(* Logix 5000 project; controller TFF vendor 1 type 14 code 107 rev 33.11; software revision 33.04; part 32 of 38 *)
(* tags used below, declared in another part *)
   ModbusLogTimer : TIMER;
   TIME : DINT[2];
   TimeInSecondsDINT : DINT;
   AI101 : ALIAS FOR AnalogPoint[16];
   AI202 : ALIAS FOR AnalogPoint[9];
   AP008 : ALIAS FOR DigitalOutput[14];
   ARC_AI101 : ARC_pH;
   ARC_AI202 : ARC_pH;
   BagInflate : BagInflate;
   DPAlarm : ALIAS FOR AlarmAnalog[40];
   FlowPath : FlowPath[64];   // Flow Path Array
   GWModbus : IO_Station;   // Status of Gateway Modbus
   IBA001 : ALIAS FOR DigitalOutput[25];
   Membrane_Data : Membrane_Data;   // Membrane Data
   ModbusTimeSyncTimer : TIMER;
   OperatingTime : OperatingTime;
   Options : Options;   // Options List
   Phase0 : ALIAS FOR Phase[0];   // Phase 0
   PI601 : ALIAS FOR AnalogPoint[21];
   PipeAnimation : PipeAnimation;   // HMI Pipe Animation Array
   SIC001_AO : ALIAS FOR AnalogOutput[0];
   SIC001_DO : ALIAS FOR DigitalOutput[8];
   SIC002_AO : ALIAS FOR AnalogOutput[1];
   SIC002_DO : ALIAS FOR DigitalOutput[9];
   SysControl : SysControl;   // General system status and command
   TimerControl : TimerControl;   // Timer Control
   TMPAlarm : ALIAS FOR AlarmAnalog[41];
   YA41 : ALIAS FOR DigitalPoint[73];
(* Process, continued *)

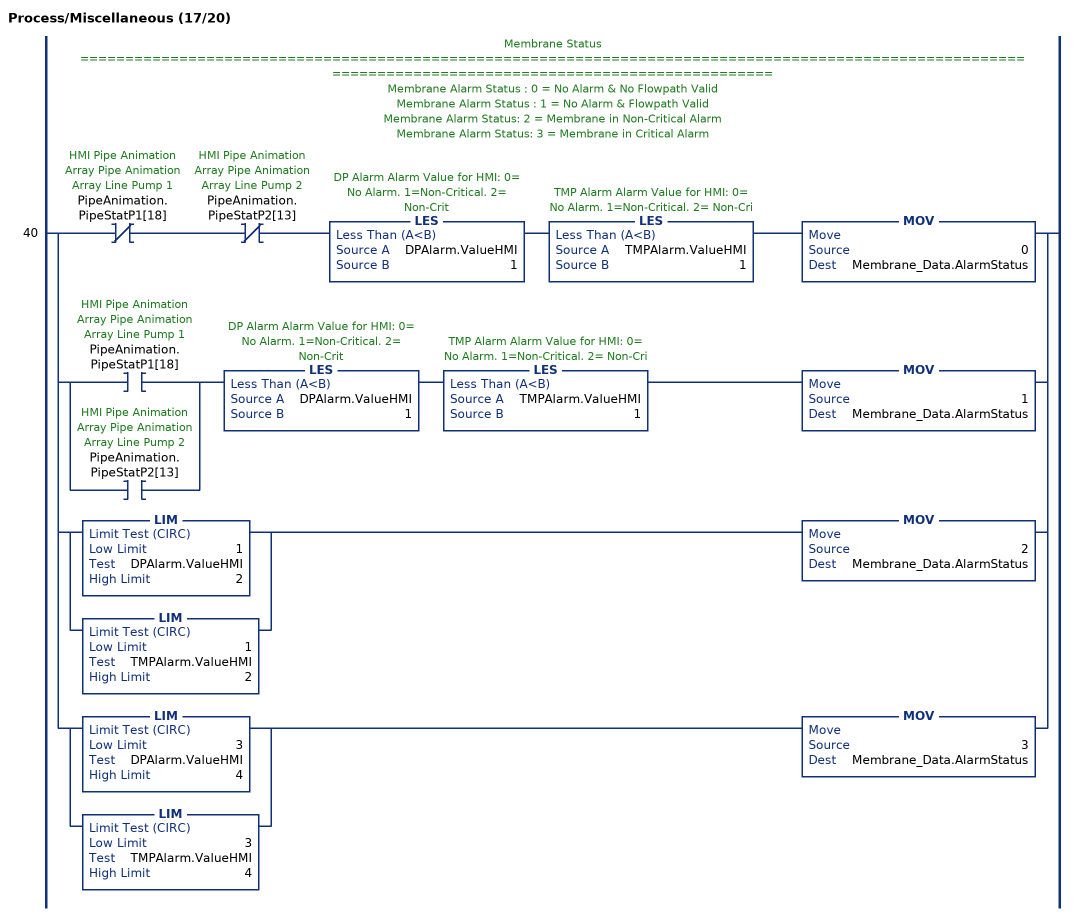
   [picture p374: Process/Miscellaneous rungs 40-40]
   // Membrane Status
   // ==========================================================================================================================================================
   // Membrane Alarm Status : 0 = No Alarm & No Flowpath Valid
   // Membrane Alarm Status : 1 = No Alarm & Flowpath Valid
   // Membrane Alarm Status: 2 = Membrane in Non-Critical Alarm
   // Membrane Alarm Status: 3 = Membrane in Critical Alarm
   40: [XIO(PipeAnimation.PipeStatP1[18]) XIO(PipeAnimation.PipeStatP2[13]) LES(DPAlarm.ValueHMI,1) LES(TMPAlarm.ValueHMI,1) MOV(0,Membrane_Data.AlarmStatus) ,[XIC(PipeAnimation.PipeStatP1[18]) ,XIC(PipeAnimation.PipeStatP2[13]) ] LES(DPAlarm.ValueHMI,1) LES(TMPAlarm.ValueHMI,1) MOV(1,Membrane_Data.AlarmStatus) ,[LIM(1,DPAlarm.ValueHMI,2) ,LIM(1,TMPAlarm.ValueHMI,2) ] MOV(2,Membrane_Data.AlarmStatus) ,[LIM(3,DPAlarm.ValueHMI,4) ,LIM(3,TMPAlarm.ValueHMI,4) ] MOV(3,Membrane_Data.AlarmStatus) ];
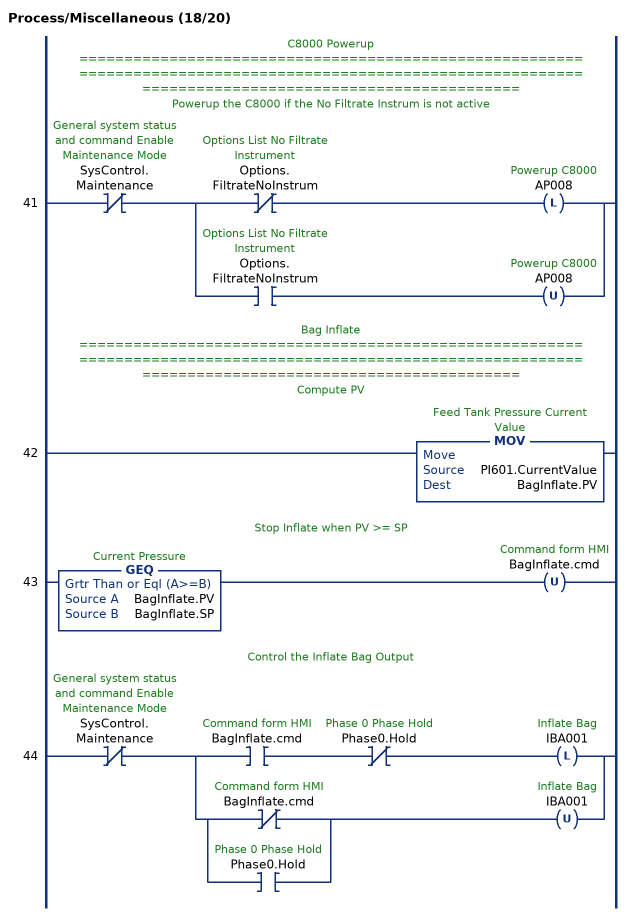
   // C8000 Powerup
   // ==========================================================================================================================================================
   // Powerup the C8000 if the No Filtrate Instrum is not active
   41: XIO(SysControl.Maintenance)[XIO(Options.FiltrateNoInstrum) OTL(AP008) ,XIC(Options.FiltrateNoInstrum) OTU(AP008) ];
   // Bag Inflate
   // ==========================================================================================================================================================
   // Compute PV
   42: MOV(PI601.CurrentValue,BagInflate.PV);
   // Stop Inflate when PV >= SP
   43: GEQ(BagInflate.PV,BagInflate.SP)OTU(BagInflate.cmd);
   // Control the Inflate Bag Output
   44: XIO(SysControl.Maintenance)[XIC(BagInflate.cmd) XIO(Phase0.Hold) OTL(IBA001) ,[XIO(BagInflate.cmd) ,XIC(Phase0.Hold) ] OTU(IBA001) ];
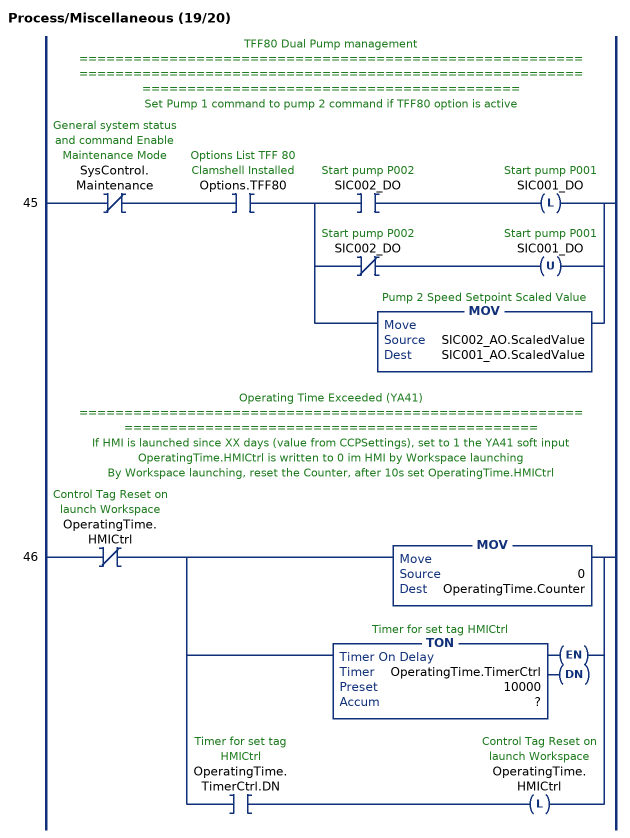
   // TFF80 Dual Pump management
   // ==========================================================================================================================================================
   // Set Pump 1 command to pump 2 command if TFF80 option is active
   45: XIO(SysControl.Maintenance)XIC(Options.TFF80)[[XIC(SIC002_DO) OTL(SIC001_DO) ,XIO(SIC002_DO) OTU(SIC001_DO) ] ,MOV(SIC002_AO.ScaledValue,SIC001_AO.ScaledValue) ];
   // Operating Time Exceeded (YA41)
   // ======================================================================================================
   // If HMI is launched since XX days (value from CCPSettings), set to 1 the YA41 soft input
   // OperatingTime.HMICtrl is written to 0 im HMI by Workspace launching
   // By Workspace launching, reset the Counter, after 10s set OperatingTime.HMICtrl
   46: XIO(OperatingTime.HMICtrl)[MOV(0,OperatingTime.Counter) ,TON(OperatingTime.TimerCtrl,?,?) ,XIC(OperatingTime.TimerCtrl.DN) OTL(OperatingTime.HMICtrl) ];
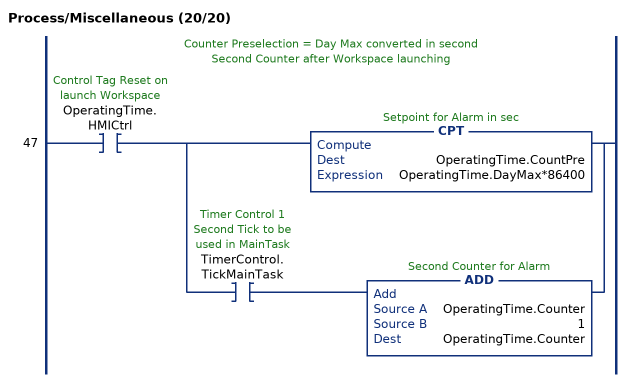
   // Counter Preselection = Day Max converted in second
   // Second Counter after Workspace launching
   47: XIC(OperatingTime.HMICtrl)[CPT(OperatingTime.CountPre,OperatingTime.DayMax*86400) ,XIC(TimerControl.TickMainTask) ADD(OperatingTime.Counter,1,OperatingTime.Counter) ];
END_ROUTINE

ROUTINE ModbusGateway   (* ladder *)
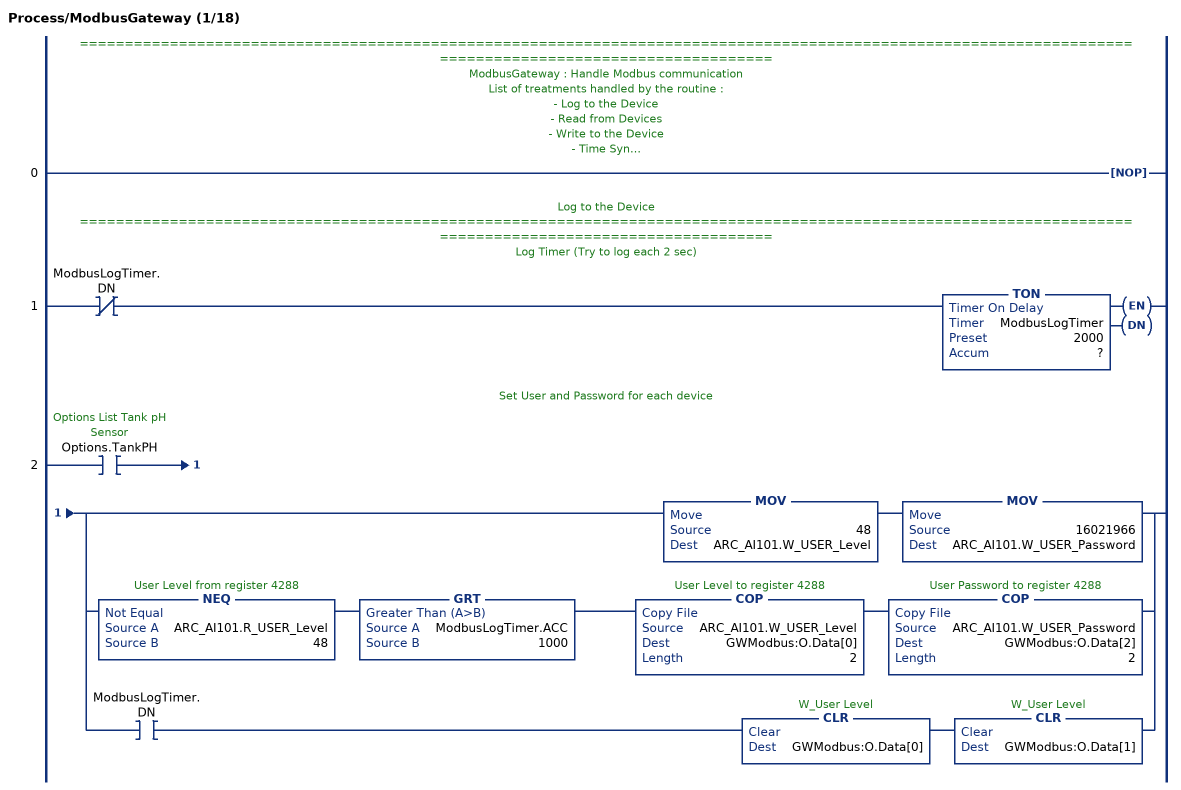
   // ==========================================================================================================================================================
   //                                                                                                                                 ModbusGateway : Handle Modbus communication
   //                                                     List of treatments handled by the routine :
   //                                                         - Log to the Device
   //                                                          - Read from Devices
   //                                                          - Write to the Device
   //                                                        - Time Sync
   //                                                     -----------------------------------------------------------------------------------------------------------------------------------------------------
   //                                                     History
   // 		2019-DEC-24 - Merck - Q. Spindler - Initial version for Candidate Release 1.00.00.00.a
   // ==========================================================================================================================================================
   0: NOP();
   // Log to the Device
   // ==========================================================================================================================================================
   // Log Timer (Try to log each 2 sec)
   1: XIO(ModbusLogTimer.DN)TON(ModbusLogTimer,?,?);
   // Set User and Password for each device
   2: XIC(Options.TankPH)[MOV(48,ARC_AI101.W_USER_Level) MOV(16021966,ARC_AI101.W_USER_Password) ,NEQ(ARC_AI101.R_USER_Level,48) GRT(ModbusLogTimer.ACC,1000) COP(ARC_AI101.W_USER_Level,GWModbus:O.Data[0],2) COP(ARC_AI101.W_USER_Password,GWModbus:O.Data[2],2) ,XIC(ModbusLogTimer.DN) CLR(GWModbus:O.Data[0]) CLR(GWModbus:O.Data[1]) ];
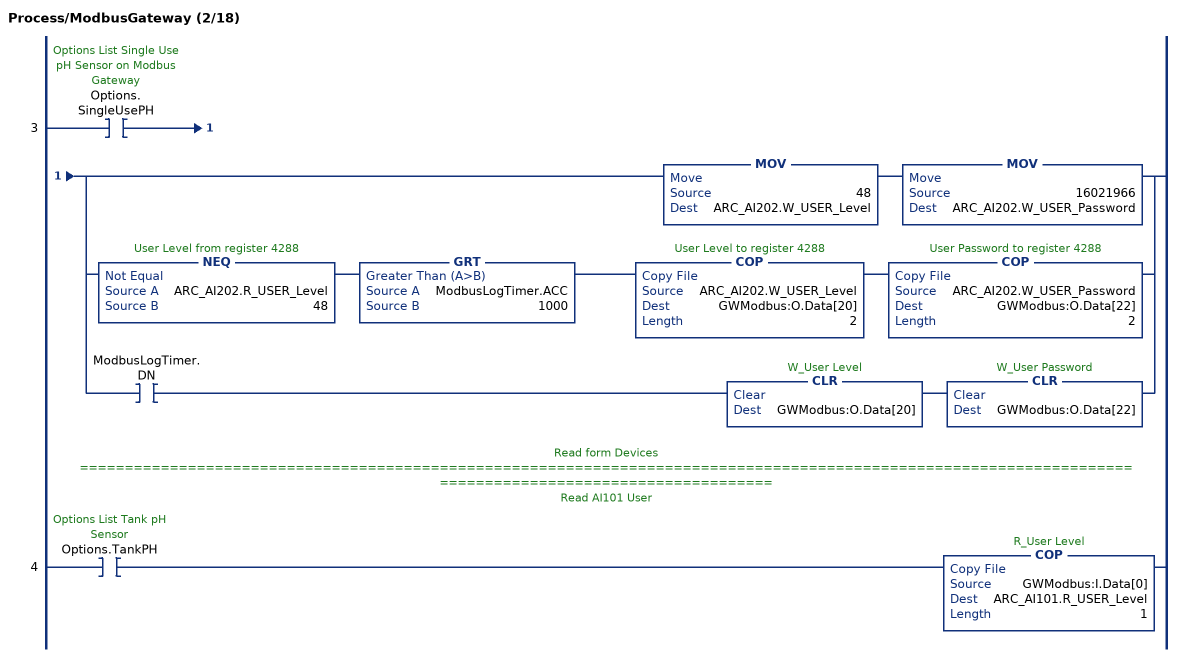
   3: XIC(Options.SingleUsePH)[MOV(48,ARC_AI202.W_USER_Level) MOV(16021966,ARC_AI202.W_USER_Password) ,NEQ(ARC_AI202.R_USER_Level,48) GRT(ModbusLogTimer.ACC,1000) COP(ARC_AI202.W_USER_Level,GWModbus:O.Data[20],2) COP(ARC_AI202.W_USER_Password,GWModbus:O.Data[22],2) ,XIC(ModbusLogTimer.DN) CLR(GWModbus:O.Data[20]) CLR(GWModbus:O.Data[22]) ];
   // Read form Devices
   // ==========================================================================================================================================================
   // Read AI101 User
   4: XIC(Options.TankPH)COP(GWModbus:I.Data[0],ARC_AI101.R_USER_Level,1);
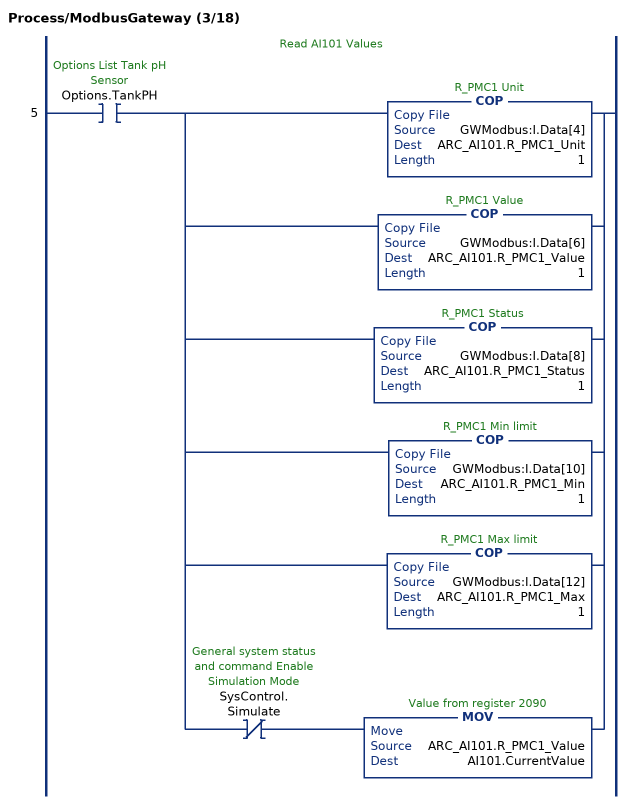
   // Read AI101 Values
   5: XIC(Options.TankPH)[COP(GWModbus:I.Data[4],ARC_AI101.R_PMC1_Unit,1) ,COP(GWModbus:I.Data[6],ARC_AI101.R_PMC1_Value,1) ,COP(GWModbus:I.Data[8],ARC_AI101.R_PMC1_Status,1) ,COP(GWModbus:I.Data[10],ARC_AI101.R_PMC1_Min,1) ,COP(GWModbus:I.Data[12],ARC_AI101.R_PMC1_Max,1) ,XIO(SysControl.Simulate) MOV(ARC_AI101.R_PMC1_Value,AI101.CurrentValue) ];
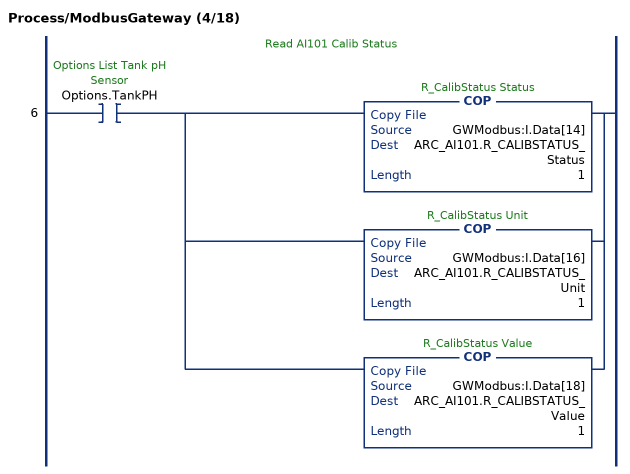
   // Read AI101 Calib Status
   6: XIC(Options.TankPH)[COP(GWModbus:I.Data[14],ARC_AI101.R_CALIBSTATUS_Status,1) ,COP(GWModbus:I.Data[16],ARC_AI101.R_CALIBSTATUS_Unit,1) ,COP(GWModbus:I.Data[18],ARC_AI101.R_CALIBSTATUS_Value,1) ];
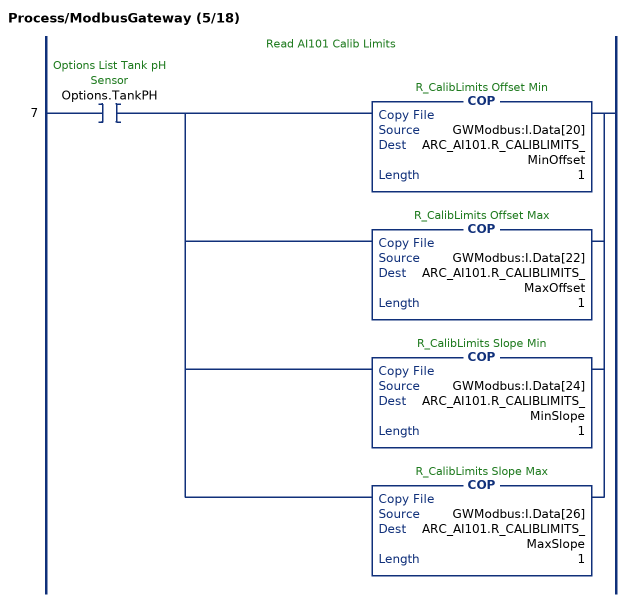
   // Read AI101 Calib Limits
   7: XIC(Options.TankPH)[COP(GWModbus:I.Data[20],ARC_AI101.R_CALIBLIMITS_MinOffset,1) ,COP(GWModbus:I.Data[22],ARC_AI101.R_CALIBLIMITS_MaxOffset,1) ,COP(GWModbus:I.Data[24],ARC_AI101.R_CALIBLIMITS_MinSlope,1) ,COP(GWModbus:I.Data[26],ARC_AI101.R_CALIBLIMITS_MaxSlope,1) ];
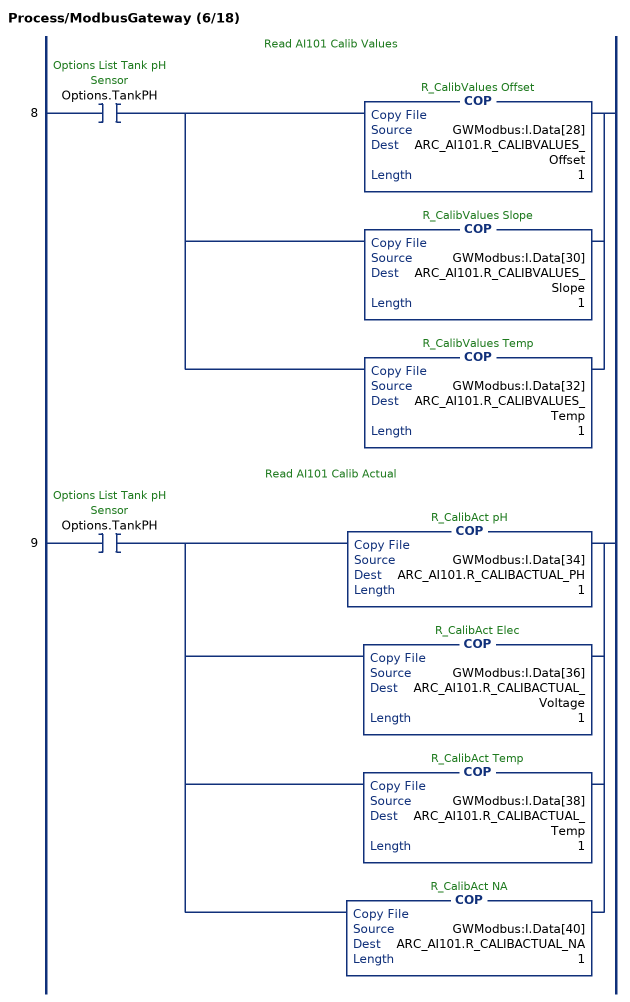
   // Read AI101 Calib Values
   8: XIC(Options.TankPH)[COP(GWModbus:I.Data[28],ARC_AI101.R_CALIBVALUES_Offset,1) ,COP(GWModbus:I.Data[30],ARC_AI101.R_CALIBVALUES_Slope,1) ,COP(GWModbus:I.Data[32],ARC_AI101.R_CALIBVALUES_Temp,1) ];
   // Read AI101 Calib Actual
   9: XIC(Options.TankPH)[COP(GWModbus:I.Data[34],ARC_AI101.R_CALIBACTUAL_PH,1) ,COP(GWModbus:I.Data[36],ARC_AI101.R_CALIBACTUAL_Voltage,1) ,COP(GWModbus:I.Data[38],ARC_AI101.R_CALIBACTUAL_Temp,1) ,COP(GWModbus:I.Data[40],ARC_AI101.R_CALIBACTUAL_NA,1) ];
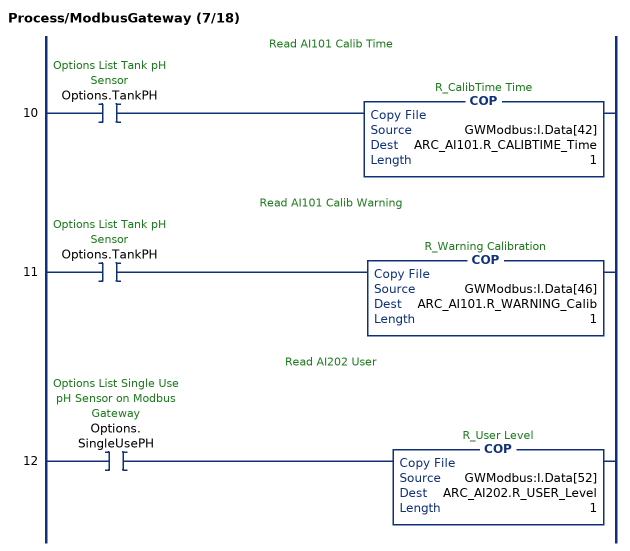
   // Read AI101 Calib Time
   10: XIC(Options.TankPH)COP(GWModbus:I.Data[42],ARC_AI101.R_CALIBTIME_Time,1);
   // Read AI101 Calib Warning
   11: XIC(Options.TankPH)COP(GWModbus:I.Data[46],ARC_AI101.R_WARNING_Calib,1);
   // Read AI202 User
   12: XIC(Options.SingleUsePH)COP(GWModbus:I.Data[52],ARC_AI202.R_USER_Level,1);
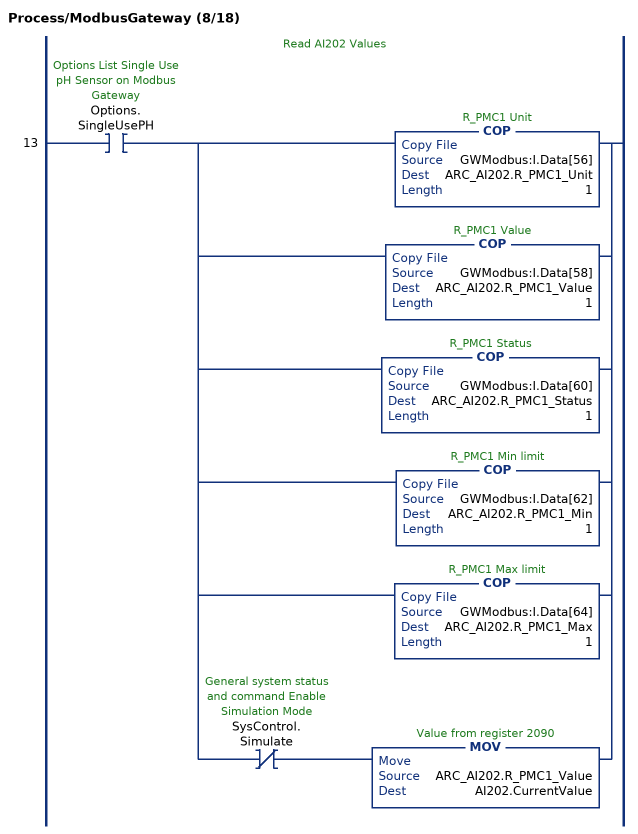
   // Read AI202 Values
   13: XIC(Options.SingleUsePH)[COP(GWModbus:I.Data[56],ARC_AI202.R_PMC1_Unit,1) ,COP(GWModbus:I.Data[58],ARC_AI202.R_PMC1_Value,1) ,COP(GWModbus:I.Data[60],ARC_AI202.R_PMC1_Status,1) ,COP(GWModbus:I.Data[62],ARC_AI202.R_PMC1_Min,1) ,COP(GWModbus:I.Data[64],ARC_AI202.R_PMC1_Max,1) ,XIO(SysControl.Simulate) MOV(ARC_AI202.R_PMC1_Value,AI202.CurrentValue) ];
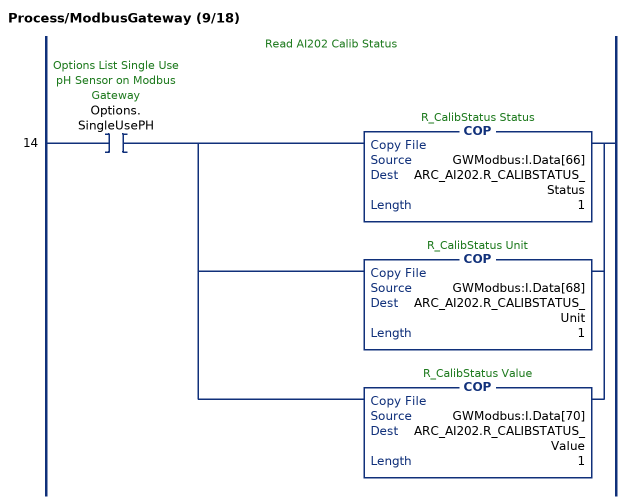
   // Read AI202 Calib Status
   14: XIC(Options.SingleUsePH)[COP(GWModbus:I.Data[66],ARC_AI202.R_CALIBSTATUS_Status,1) ,COP(GWModbus:I.Data[68],ARC_AI202.R_CALIBSTATUS_Unit,1) ,COP(GWModbus:I.Data[70],ARC_AI202.R_CALIBSTATUS_Value,1) ];
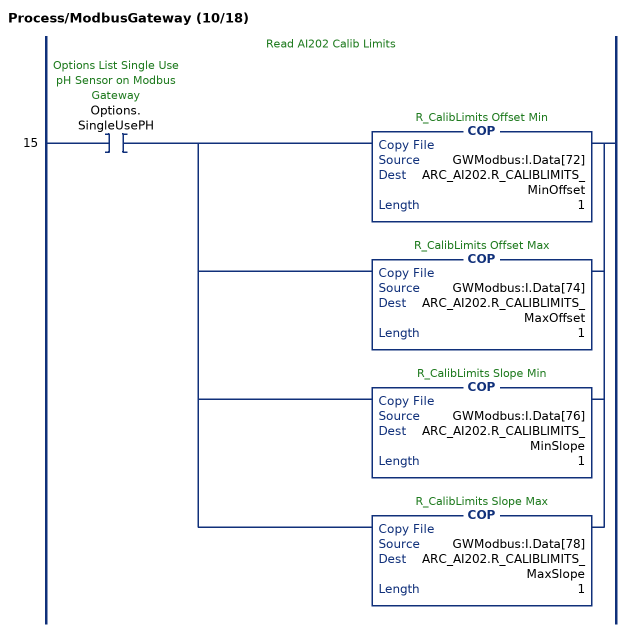
   // Read AI202 Calib Limits
   15: XIC(Options.SingleUsePH)[COP(GWModbus:I.Data[72],ARC_AI202.R_CALIBLIMITS_MinOffset,1) ,COP(GWModbus:I.Data[74],ARC_AI202.R_CALIBLIMITS_MaxOffset,1) ,COP(GWModbus:I.Data[76],ARC_AI202.R_CALIBLIMITS_MinSlope,1) ,COP(GWModbus:I.Data[78],ARC_AI202.R_CALIBLIMITS_MaxSlope,1) ];
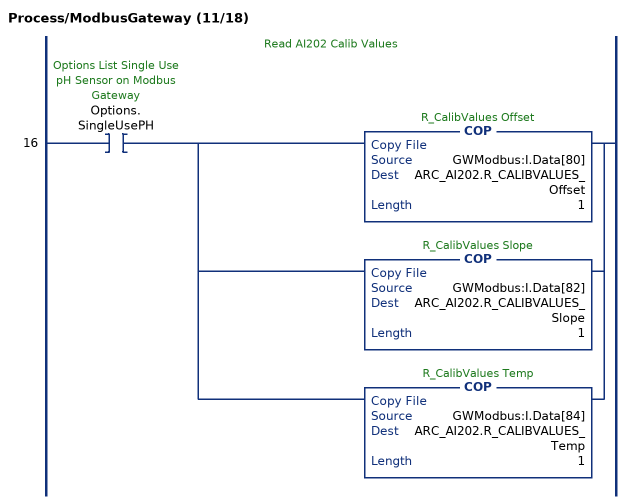
   // Read AI202 Calib Values
   16: XIC(Options.SingleUsePH)[COP(GWModbus:I.Data[80],ARC_AI202.R_CALIBVALUES_Offset,1) ,COP(GWModbus:I.Data[82],ARC_AI202.R_CALIBVALUES_Slope,1) ,COP(GWModbus:I.Data[84],ARC_AI202.R_CALIBVALUES_Temp,1) ];
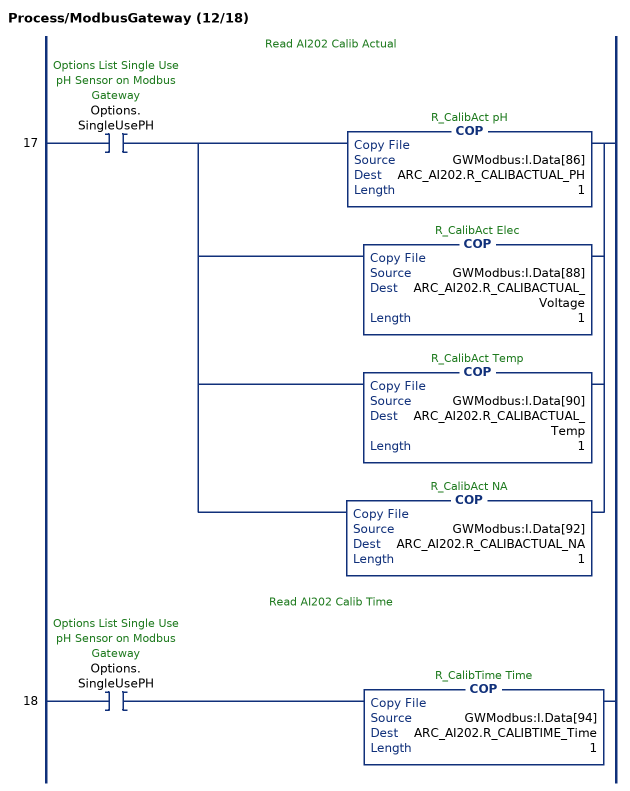
   // Read AI202 Calib Actual
   17: XIC(Options.SingleUsePH)[COP(GWModbus:I.Data[86],ARC_AI202.R_CALIBACTUAL_PH,1) ,COP(GWModbus:I.Data[88],ARC_AI202.R_CALIBACTUAL_Voltage,1) ,COP(GWModbus:I.Data[90],ARC_AI202.R_CALIBACTUAL_Temp,1) ,COP(GWModbus:I.Data[92],ARC_AI202.R_CALIBACTUAL_NA,1) ];
   // Read AI202 Calib Time
   18: XIC(Options.SingleUsePH)COP(GWModbus:I.Data[94],ARC_AI202.R_CALIBTIME_Time,1);
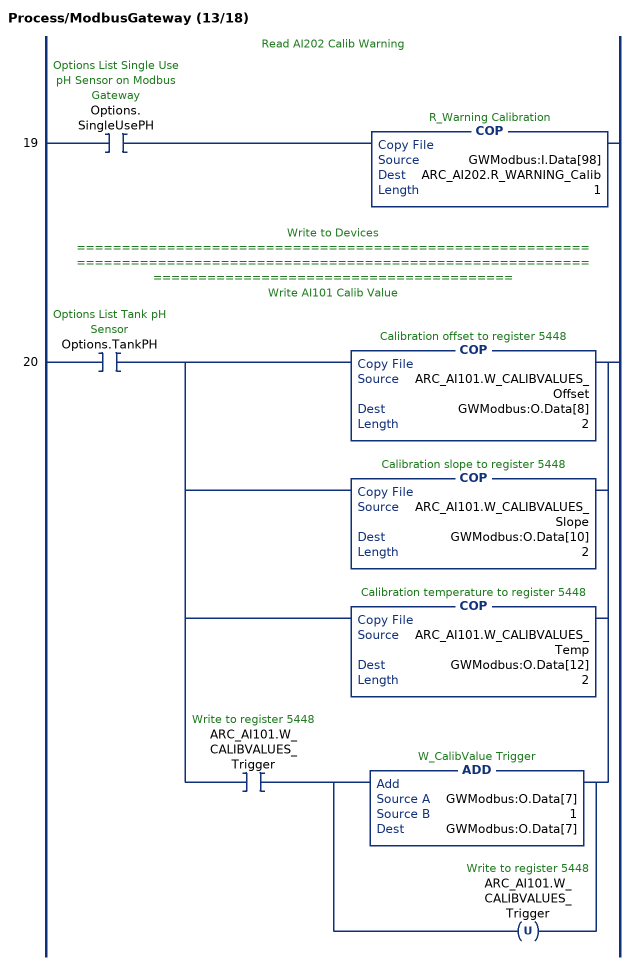
   // Read AI202 Calib Warning
   19: XIC(Options.SingleUsePH)COP(GWModbus:I.Data[98],ARC_AI202.R_WARNING_Calib,1);
   // Write to Devices
   // ==========================================================================================================================================================
   // Write AI101 Calib Value
   20: XIC(Options.TankPH)[COP(ARC_AI101.W_CALIBVALUES_Offset,GWModbus:O.Data[8],2) ,COP(ARC_AI101.W_CALIBVALUES_Slope,GWModbus:O.Data[10],2) ,COP(ARC_AI101.W_CALIBVALUES_Temp,GWModbus:O.Data[12],2) ,XIC(ARC_AI101.W_CALIBVALUES_Trigger) [ADD(GWModbus:O.Data[7],1,GWModbus:O.Data[7]) ,OTU(ARC_AI101.W_CALIBVALUES_Trigger) ] ];
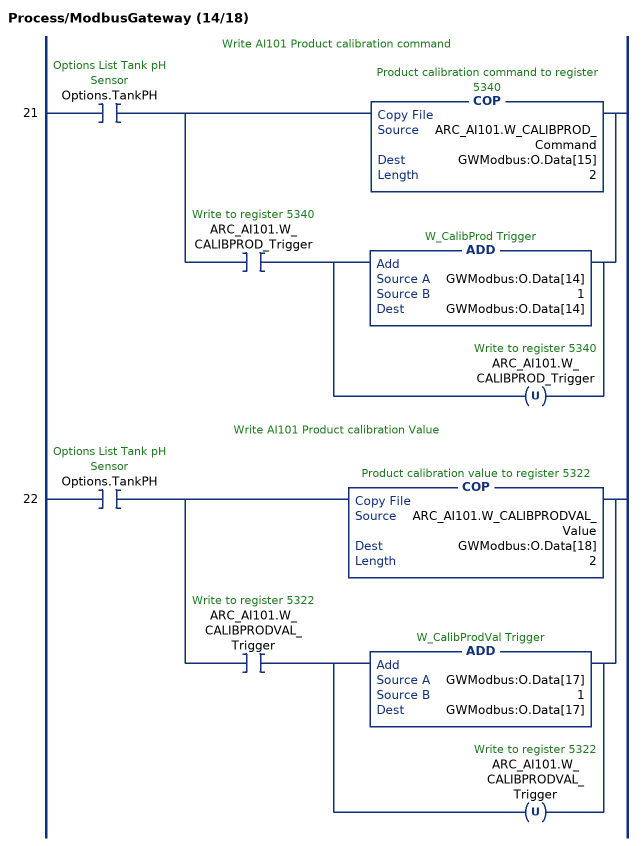
   // Write AI101 Product calibration command
   21: XIC(Options.TankPH)[COP(ARC_AI101.W_CALIBPROD_Command,GWModbus:O.Data[15],2) ,XIC(ARC_AI101.W_CALIBPROD_Trigger) [ADD(GWModbus:O.Data[14],1,GWModbus:O.Data[14]) ,OTU(ARC_AI101.W_CALIBPROD_Trigger) ] ];
   // Write AI101 Product calibration Value
   22: XIC(Options.TankPH)[COP(ARC_AI101.W_CALIBPRODVAL_Value,GWModbus:O.Data[18],2) ,XIC(ARC_AI101.W_CALIBPRODVAL_Trigger) [ADD(GWModbus:O.Data[17],1,GWModbus:O.Data[17]) ,OTU(ARC_AI101.W_CALIBPRODVAL_Trigger) ] ];
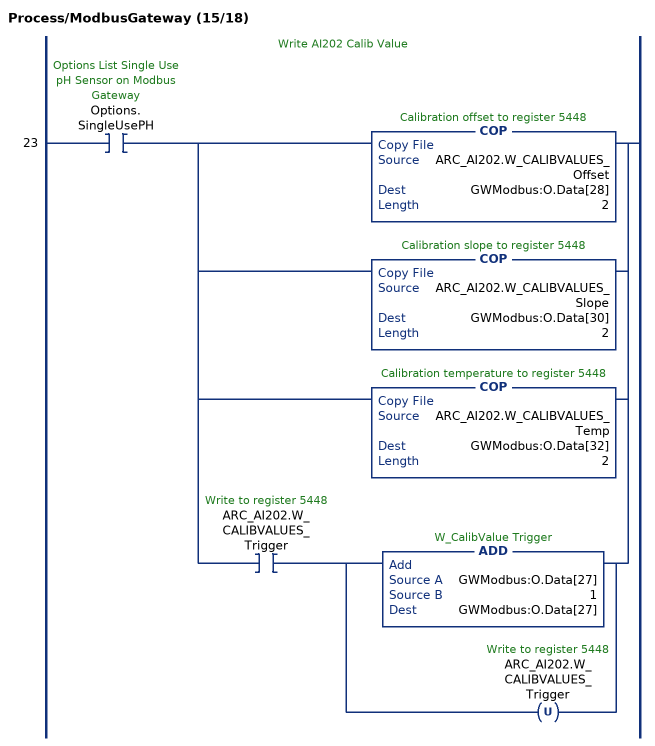
   // Write AI202 Calib Value
   23: XIC(Options.SingleUsePH)[COP(ARC_AI202.W_CALIBVALUES_Offset,GWModbus:O.Data[28],2) ,COP(ARC_AI202.W_CALIBVALUES_Slope,GWModbus:O.Data[30],2) ,COP(ARC_AI202.W_CALIBVALUES_Temp,GWModbus:O.Data[32],2) ,XIC(ARC_AI202.W_CALIBVALUES_Trigger) [ADD(GWModbus:O.Data[27],1,GWModbus:O.Data[27]) ,OTU(ARC_AI202.W_CALIBVALUES_Trigger) ] ];
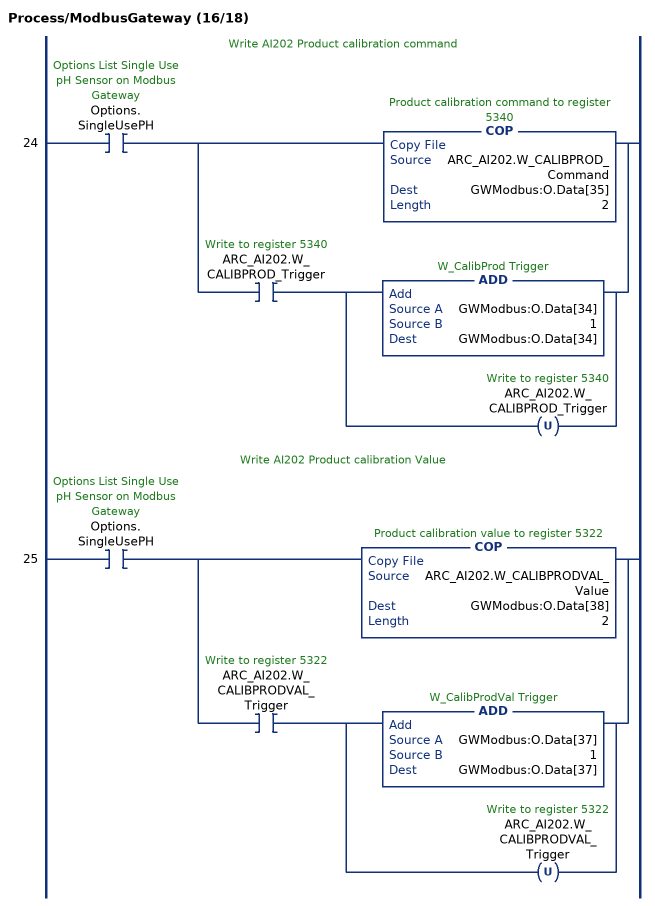
   // Write AI202 Product calibration command
   24: XIC(Options.SingleUsePH)[COP(ARC_AI202.W_CALIBPROD_Command,GWModbus:O.Data[35],2) ,XIC(ARC_AI202.W_CALIBPROD_Trigger) [ADD(GWModbus:O.Data[34],1,GWModbus:O.Data[34]) ,OTU(ARC_AI202.W_CALIBPROD_Trigger) ] ];
   // Write AI202 Product calibration Value
   25: XIC(Options.SingleUsePH)[COP(ARC_AI202.W_CALIBPRODVAL_Value,GWModbus:O.Data[38],2) ,XIC(ARC_AI202.W_CALIBPRODVAL_Trigger) [ADD(GWModbus:O.Data[37],1,GWModbus:O.Data[37]) ,OTU(ARC_AI202.W_CALIBPRODVAL_Trigger) ] ];
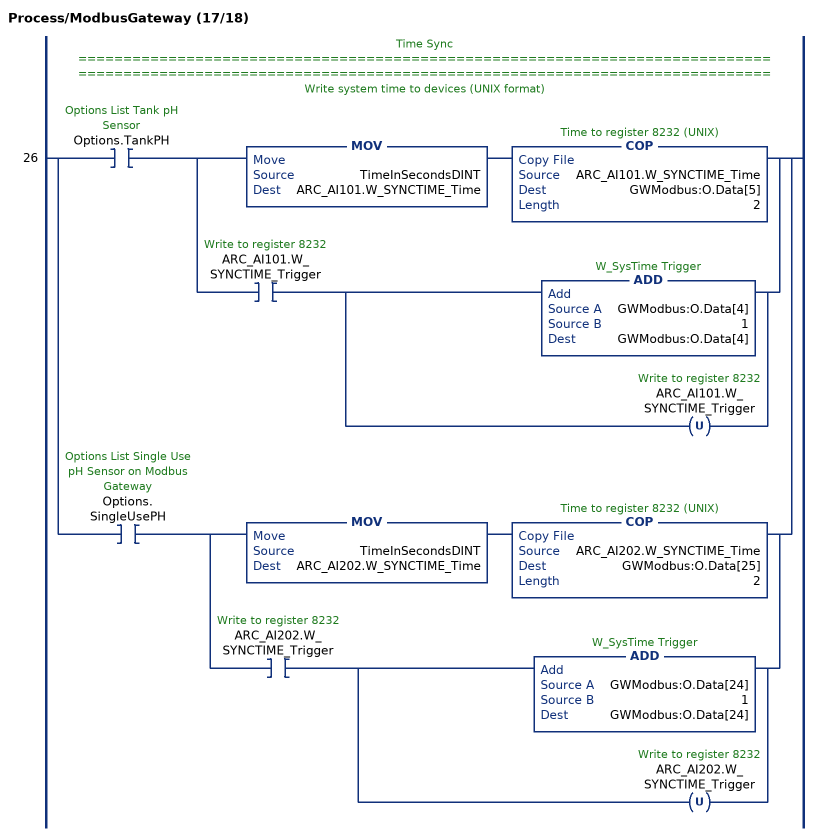
   // Time Sync
   // ==========================================================================================================================================================
   // Write system time to devices (UNIX format)
   26: [XIC(Options.TankPH) [MOV(TimeInSecondsDINT,ARC_AI101.W_SYNCTIME_Time) COP(ARC_AI101.W_SYNCTIME_Time,GWModbus:O.Data[5],2) ,XIC(ARC_AI101.W_SYNCTIME_Trigger) [ADD(GWModbus:O.Data[4],1,GWModbus:O.Data[4]) ,OTU(ARC_AI101.W_SYNCTIME_Trigger) ] ] ,XIC(Options.SingleUsePH) [MOV(TimeInSecondsDINT,ARC_AI202.W_SYNCTIME_Time) COP(ARC_AI202.W_SYNCTIME_Time,GWModbus:O.Data[25],2) ,XIC(ARC_AI202.W_SYNCTIME_Trigger) [ADD(GWModbus:O.Data[24],1,GWModbus:O.Data[24]) ,OTU(ARC_AI202.W_SYNCTIME_Trigger) ] ] ];
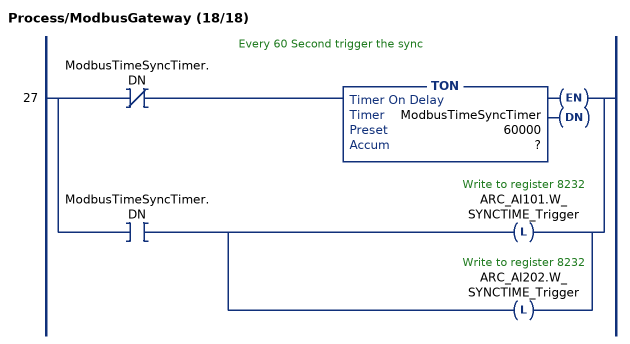
   // Every 60 Second trigger the sync
   27: [XIO(ModbusTimeSyncTimer.DN) TON(ModbusTimeSyncTimer,?,?) ,XIC(ModbusTimeSyncTimer.DN) [OTL(ARC_AI101.W_SYNCTIME_Trigger) ,OTL(ARC_AI202.W_SYNCTIME_Trigger) ] ];
END_ROUTINE
